(* PLC project g_door_reversal_momentary, Anonymous Benchmark Suite 1.0 *)
(* stored: creationDateTime 2026-08-28T00:00:00 *)

PROGRAM g_door_reversal_momentary
  VAR_INPUT
    CloseCmd : BOOL;
    OpenCmd : BOOL;
    Beam : BOOL;
    TopLimit : BOOL;
  END_VAR
  VAR_OUTPUT
    Reversing : BOOL;
    MoveDown : BOOL;
    MoveUp : BOOL;
  END_VAR

(* LD diagram, written out as Structured Text *)
Reversing := Beam AND NOT TopLimit;
MoveDown := CloseCmd AND NOT Beam AND NOT Reversing;
MoveUp := OpenCmd OR Reversing;
END_PROGRAM

CONFIGURATION Config0
  RESOURCE Res0 ON PLC
    TASK tcyclic(INTERVAL := T#10ms, PRIORITY := 0);
    PROGRAM inst0 WITH tcyclic : g_door_reversal_momentary;
  END_RESOURCE
END_CONFIGURATION
